# EPICS autosave request: iocs/quadem/ah401-ioc/auto_settings.req
file "quadEM_IOC_settings.req",        P=$(P), R=$(R)
